// TIA Portal V20 export
Screen "Pop-up_Sealer_2"  395x650
  ScreenItem "Robot Name" at 2,2 size 393x48  Type=HmiIOField
  ScreenItem "Background" at 2,48 size 393x602  Type=HmiRectangle
  ScreenItem "Cancel Mode" at 315,4 size 76x42  Type=HmiButton
  ScreenItem "矩形_4" at 36,76 size 324x517  Type=HmiRectangle
  ScreenItem "Text Filed E- Stop_17" at 44,341 size 148x21  Type=HmiTextBox
  ScreenItem "Text Field In Auto On_9" at 44,106 size 148x21  Type=HmiTextBox
  ScreenItem "Text Field Home Position_17" at 44,129 size 148x21  Type=HmiTextBox
  ScreenItem "Text field Robot Status_5" at 36,77 size 324x26  Type=HmiTextBox
  ScreenItem "Text Field Manual_17" at 44,271 size 148x21  Type=HmiTextBox
  ScreenItem "Text Field System Ready_9" at 44,153 size 148x21  Type=HmiTextBox
  ScreenItem "Text Field Motor On_9" at 44,176 size 148x21  Type=HmiTextBox
  ScreenItem "Text Field In Cycle_9" at 44,200 size 148x21  Type=HmiTextBox
  ScreenItem "Text Field Cycle On_17" at 44,223 size 148x21  Type=HmiTextBox
  ScreenItem "Text Field On Path_17" at 44,247 size 148x21  Type=HmiTextBox
  ScreenItem "Text Field Tryout Mode_17" at 44,294 size 148x21  Type=HmiTextBox
  ScreenItem "Text Field Stop_17" at 44,318 size 148x21  Type=HmiTextBox
  ScreenItem "Text Filed Error_9" at 44,365 size 148x21  Type=HmiTextBox
  ScreenItem "Text Filed Process Fault_9" at 44,388 size 148x21  Type=HmiTextBox
  ScreenItem "Text Field Home Position_18" at 44,412 size 148x21  Type=HmiTextBox
  ScreenItem "Text Filed E- Stop_18" at 44,554 size 148x21  Type=HmiTextBox
  ScreenItem "Text Field Manual_18" at 44,483 size 148x21  Type=HmiTextBox
  ScreenItem "Text Field Cycle On_18" at 44,436 size 148x21  Type=HmiTextBox
  ScreenItem "Text Field On Path_18" at 44,459 size 148x21  Type=HmiTextBox
  ScreenItem "Text Field Tryout Mode_18" at 44,506 size 148x21  Type=HmiTextBox
  ScreenItem "Text Field Stop_18" at 44,530 size 148x21  Type=HmiTextBox
  ScreenItem "Text Filed E- Stop_19" at 205,341 size 148x21  Type=HmiTextBox
  ScreenItem "Text Field In Auto On_10" at 205,106 size 148x21  Type=HmiTextBox
  ScreenItem "Text Field Home Position_19" at 205,129 size 148x21  Type=HmiTextBox
  ScreenItem "Text Field Manual_19" at 205,271 size 148x21  Type=HmiTextBox
  ScreenItem "Text Field System Ready_10" at 205,153 size 148x21  Type=HmiTextBox
  ScreenItem "Text Field Motor On_10" at 205,176 size 148x21  Type=HmiTextBox
  ScreenItem "Text Field In Cycle_10" at 205,200 size 148x21  Type=HmiTextBox
  ScreenItem "Text Field Cycle On_19" at 205,223 size 148x21  Type=HmiTextBox
  ScreenItem "Text Field On Path_19" at 205,247 size 148x21  Type=HmiTextBox
  ScreenItem "Text Field Tryout Mode_19" at 205,294 size 148x21  Type=HmiTextBox
  ScreenItem "Text Field Stop_19" at 205,318 size 148x21  Type=HmiTextBox
  ScreenItem "Text Filed Error_10" at 205,365 size 148x21  Type=HmiTextBox
  ScreenItem "Text Filed Process Fault_10" at 205,388 size 148x21  Type=HmiTextBox
  ScreenItem "Text Field Home Position_20" at 205,412 size 148x21  Type=HmiTextBox
  ScreenItem "Text Filed E- Stop_20" at 205,554 size 148x21  Type=HmiTextBox
  ScreenItem "Text Field Manual_20" at 205,483 size 148x21  Type=HmiTextBox
  ScreenItem "Text Field Cycle On_20" at 205,436 size 148x21  Type=HmiTextBox
  ScreenItem "Text Field On Path_20" at 205,459 size 148x21  Type=HmiTextBox
  ScreenItem "Text Field Tryout Mode_20" at 205,506 size 148x21  Type=HmiTextBox
  ScreenItem "Text Field Stop_20" at 205,530 size 148x21  Type=HmiTextBox
